FUNCTION_BLOCK fb_Dev_Actuator EXTENDS abs_fb_Device
VAR_INPUT
	IO_Input_Feedback : BOOL;
END_VAR

VAR_IN_OUT
	IO_Output_Actuate : BOOL;
END_VAR

VAR
	HMI						: ST_Actuator_HMI_Interface;
	_setActuate 			: BOOL;
	_retractOnFault			: BOOL;
	_hasFeedback			: BOOL;
	_faultH_onDelay			: TON;
	_faultH_offDelay		: TON;
	_faultH_OnDelay_Trigger	: BOOL;
	_faultH_OffDelay_Trigger: BOOL;
	_onDelay_time			: TIME;
	_offDelay_time			: TIME;
	_InvFeedback			: BOOL;
	_actuatorFeedback		: BOOL;
	_maintainAutoState		: BOOL;
	_disableHMIControl		: BOOL;
END_VAR

VAR_OUTPUT
	stsActuated : BOOL;

END_VAR

DeviceLogic();
Interlock.name := _DeviceName;
Interlock(inpConfig := _dataInterlock);

// Flip feedback if cofigured for inverted feedback
IF _InvFeedback THEN
	IF IO_Input_Feedback THEN
		_actuatorFeedback := FALSE;
	ELSE
		_actuatorFeedback :=TRUE;
	END_IF
ELSE
	IF IO_Input_Feedback THEN
		_actuatorFeedback :=TRUE;
	ELSE
		_actuatorFeedback :=FALSE;
	END_IF
END_IF

// If no IO based feedback, set actuation state for feedback
IF _hasFeedback THEN
	stsActuated := _actuatorFeedback;
ELSE
	stsActuated := _setActuate;
END_IF

// Check for timeouts
FaultHandler(_actuatorFeedback);

// Control via HMI if in manual
// cmdActuate an cmdRetract methods only work in Auto, unless
// device is configured for no manual control
IF NOT _disableHMIControl THEN
	IF NOT _inAuto THEN 
		IF HMI.ocmdActuate THEN
			cmdActuate();
		ELSE
			cmdRetract();
		END_IF
	ELSE
		// if property set, change the HMI actuatoion toggle state so that
		// transition from auto to manual does not change the state
		// otherwise upon transition HMI will change state to whatever it was in manual last
		IF _maintainAutoState THEN
			HMI.ocmdActuate := _setActuate;
		END_IF
	END_IF
END_IF
// Configure retract on feedback
IF stsFaulted AND _retractOnFault THEN
	HMI.ocmdActuate := 0;
	_setActuate		:= 0;
END_IF

// Log state changes
IF _setActuate THEN
	IO_output_actuate :=TRUE;
	sendLog('Actuating ON',1);
ELSE
	IO_output_actuate :=FALSE;
	sendLog('Actuating OFF',1);
END_IF

HMI.HMIbaseDevice := HMIbaseDevice;
HMI.stsActuated   := stsActuated;
HMI.setActuate    := _setActuate;

PROPERTY cfgDeviceName : string
GET
cfgDeviceName := _DeviceName;
END_GET
SET
_DeviceName := cfgDeviceName;
END_SET
END_PROPERTY

PROPERTY cfgDisableHMIControl : BOOL
GET
cfgDisableHMIControl := _disableHMIControl;
END_GET
SET
_disableHMIControl := cfgDisableHMIControl;
END_SET
END_PROPERTY

PROPERTY cfgHasFeedback : BOOL
GET
cfgHasFeedback := _hasFeedback;
END_GET
SET
_hasFeedback	:= cfgHasFeedback;
END_SET
END_PROPERTY

PROPERTY PUBLIC cfgInvFeedback : Bool
GET
cfgInvFeedback := _InvFeedback;
END_GET
SET
_InvFeedback := cfgInvFeedback;
END_SET
END_PROPERTY

PROPERTY cfgMaintainAutoState : BOOL
GET
cfgMaintainAutoState	:= _maintainAutoState;
END_GET
SET
_maintainAutoState := cfgMaintainAutoState;
END_SET
END_PROPERTY

PROPERTY cfgOffDelay : TIME
GET
cfgOffDelay := _offDelay_time;
END_GET
SET
_offDelay_time := cfgOffDelay;
END_SET
END_PROPERTY

PROPERTY PUBLIC cfgOnDelay : Time
GET
cfgOnDelay := _onDelay_time;
END_GET
SET
_OnDelay_time := cfgOnDelay;
END_SET
END_PROPERTY

PROPERTY cfgRetractOnFault : bool
GET
cfgRetractOnFault := _retractOnFault;
END_GET
SET
_retractOnFault := cfgRetractOnFault;
END_SET
END_PROPERTY

METHOD PUBLIC cmdActuate : BOOL
VAR_INPUT
	
END_VAR
IF Interlock.outInterlockOK AND NOT stsFaulted THEN
	_setActuate :=TRUE;
END_IF
END_METHOD

METHOD cmdReset : BOOL
IF stsFaulted THEN
	setFault(0,'');
END_IF
END_METHOD

METHOD PUBLIC cmdRetract : BOOL
VAR_INPUT
END_VAR
// Retracting (de-energising) is always allowed. It used to require the interlock to be met,
// so an actuator whose interlock dropped could not be switched off, by the operator or by code,
// unless cfgRetractOnFault happened to be set.
_setActuate := FALSE;
END_METHOD

METHOD PRIVATE FaultHandler : BOOL
VAR_INPUT
	inpFeedback : BOOL; 
	
END_VAR
//if setActuate, set timer. If timer done and no feedback, then fault
IF (_onDelay_Time <> T#0S) AND _hasfeedback THEN
	_faultH_onDelay(IN:=_faultH_OnDelay_Trigger,PT:=_onDelay_time);
	IF (NOT stsFaulted) AND _setActuate THEN
		_faultH_OnDelay_Trigger := TRUE;
		IF _faultH_onDelay.Q AND NOT _actuatorFeedback THEN
			setFault(1,'actuator feedback missing.');
		END_IF
	ELSE
		_faultH_OnDelay_Trigger := FALSE;
	END_IF
END_IF

IF (_offDelay_Time <> T#0S) AND _hasfeedback THEN
	_faultH_offDelay(IN:=_faultH_OffDelay_Trigger,PT:=_offDelay_time);
	IF (NOT stsFaulted) AND NOT(_setActuate) THEN
		_faultH_OffDelay_Trigger := TRUE;
		IF _faultH_offDelay.Q AND _actuatorFeedback THEN
			setFault(1,'Feedback present when not actuated.');
		END_IF
	ELSE
		_faultH_OffDelay_Trigger := FALSE;
	END_IF
END_IF


//IF _actuatorFeedback AND NOT(_setActuate) and _hasFeedback THEN
//	setFault(1,'Feedback present when not actuated');
//END_IF

//if not actuated but feedback is in, actuator is stuck closed
//+TODO

//If enabled and cmdActuated and lost interlock, then fault
IF NOT stsFaulted AND _setActuate THEN
	IF NOT interlock.outInterlockOK THEN
		setFault(1,CONCAT('I_NOK - ',Interlock.stsFirstOut));
	END_IF
END_IF
END_METHOD

//FB_Init is always available implicitly and it is used primarily for initialization.
//The return value is not evaluated. For a specific influence, you can also declare the
//methods explicitly and provide additional code there with the standard initialization
//code. You can evaluate the return value.
METHOD FB_Init: BOOL
VAR_INPUT
    bInitRetains: BOOL; // TRUE: the retain variables are initialized (reset warm / reset cold)
    bInCopyCode: BOOL;  // TRUE: the instance will be copied to the copy code afterward (online change)
	
	cfgDeviceName 		: STRING;
	cfgEnable 			: BOOL;
	cfgInitEventClass	: BOOL;
	cfgOnDelay 			: TIME;
	cfgOffDelay			: TIME;
	cfgRetractOnFault 	: BOOL;
	cfgInvFeedback		: BOOL; 
	cfgHasFeedback		: BOOL;

END_VAR
THIS^.cfgDeviceName 		:= 		cfgDeviceName; 
THIS^.cfgEnable				:=		cfgEnable;
THIS^.cfgInitEventClass		:= 		cfgInitEventClass;		
THIS^.cfgOnDelay 			:= 		cfgOnDelay; 
THIS^.cfgOffDelay			:=		cfgOffDelay;			
THIS^.cfgRetractOnFault		:=      cfgRetractOnFault;
THIS^.cfgInvFeedback		:=		cfgInvFeedback;
THIS^.cfgHasFeedback		:=		cfgHasFeedback;
END_METHOD

END_FUNCTION_BLOCK

(* stored: Version 1.1.0.1
   POU fb_Dev_Actuator: Id {81e85ebb-2100-42fa-8869-8bedf307b98d}, SpecialFunc None
   Folder Privates: Id {98a5be4d-699f-42e4-a6a5-0814ff6a062c}
   Property cfgDeviceName: Id {2aba6988-1e9a-49ec-be4d-c870e6164032}
   Get Get: Id {76d50d17-8d13-4ef8-8dc2-085e0561228b}
   Set Set: Id {19205351-3140-4d8a-bea4-36b4987c7f42}
   Property cfgDisableHMIControl: Id {6a47590d-e86b-4ea1-bec8-d054a068d0f8}
   Get Get: Id {bdebbfb4-23cf-4922-81ec-81865239ed10}
   Set Set: Id {5fabe481-e236-4694-9ab9-ddb5cd0b6aae}
   Property cfgHasFeedback: Id {6e651f8c-1b21-4f4d-9868-d1ace3f1d0ca}
   Get Get: Id {c7c1390b-d4b1-4e66-8872-22ebb11d73c9}
   Set Set: Id {3a3f1ab7-e211-47e2-a854-ff9a34cbd1be}
   Property cfgInvFeedback: Id {bd80d261-bdf7-4785-97c6-05fb89928191}
   Get Get: Id {7027c690-2075-4984-8071-f53056d2d55e}
   Set Set: Id {87ed1395-350e-49c2-b5bb-18a4482f8c88}
   Property cfgMaintainAutoState: Id {6373a2c8-0ef1-491f-a176-7dd6c8964993}
   Get Get: Id {852e4d43-d893-4b31-abfb-f926ce93824f}
   Set Set: Id {0da50087-6028-4c91-8d46-307051213243}
   Property cfgOffDelay: Id {0605322d-9aa5-48dd-a138-12eb219aafbe}
   Get Get: Id {e82ca65e-b818-4216-bda5-e75bba3fef38}
   Set Set: Id {f82b13df-7f79-41ca-8253-659c448d5ac3}
   Property cfgOnDelay: Id {aab5577b-6b87-4620-9d52-95d00ea2e676}
   Get Get: Id {3de0fb61-aec3-44dc-96ac-ff138be1c7ca}
   Set Set: Id {7af5c5a3-99e4-4728-b6ab-9656302c7602}
   Property cfgRetractOnFault: Id {27f75573-9d03-472c-9d37-97a6875b6a41}
   Get Get: Id {d64de5a2-24bf-4d2c-bf67-ab41b582a9ec}
   Set Set: Id {e0248c55-875c-4cbc-9384-469b45799dad}
   Method cmdActuate: Id {0e9fda91-8d5f-4566-a5c5-acf49981b4f4}
   Method cmdReset: Id {11ab5455-1962-4f91-aeda-b84e24d3ac25}
   Method cmdRetract: Id {a721761f-2f78-4f45-88de-6492373238ef}
   Method FaultHandler: Id {a88fc260-ac03-4357-9f5c-cfcc4dfecdaf}
   Method FB_Init: Id {7407b03c-e4e5-4437-a988-6afe951e456e} *)
